(*
SPDX-FileCopyrightText: © 2026 Oleksandr Tiutyk <trofimich@gmail.com>
SPDX-License-Identifier: MIT
License: https://opensource.org/license/mit
*)

(*!
<summary>
Beckhoff bidirectional power measurement phase channel process image.
</summary>
<description>
Combines an EL3413/EL3433 phase input PDO, including mandatory Status, with its output Index selector.
Evaluate input validity and wait for In.Index to acknowledge Out.Index before interpreting In.VariantValue.
EL3403 uses EL3403_CHANNEL; its phase status flags are different. Link input/output fields individually.
Use one owner task and synchronize other access; copying stores data without creating new hardware links.
When used for I/O, link located fields or their containing buffers to the matching selected PDOs.
The record is not a packed wire buffer; compiler padding is not part of the device specification.
Unlinked/default values do not prove valid I/O. The caller evaluates bus/channel validity before use.
Use one owner task per instance and externally synchronize other access; multi-field snapshots are not atomic.
Copies store data without creating hardware links. Keep borrowed field references valid while consumers are bound.
This passive record performs no validation, synchronization, configuration or protocol advancement.
</description>
*)
TYPE POWER_MEASUREMENT_CHANNEL :
STRUCT
	In : POWER_MEASUREMENT_INPUT_CHANNEL;
	Out : POWER_MEASUREMENT_OUTPUT_CHANNEL;
END_STRUCT
END_TYPE

(* stored: Version 1.1.0.1, ProductVersion 3.1.4026.20
   DUT POWER_MEASUREMENT_CHANNEL: Id {2ca088d6-6422-4995-951b-814c1760935c} *)
